(* Logix 5000 project; controller TFF vendor 1 type 14 code 107 rev 34.11; software revision 34.03; part 30 of 36 *)
(* tags used below, declared in another part *)
   Address : DINT;   // Temp Address
   Index : DINT;   // Index
   Index2 : DINT;   // Index
   ACQ002 : ALIAS FOR DigitalOutput[0];   // Emergency Stop Acknowledge
   AlarmControl : AlarmControl;   // Alarm Control
   AnalogOutput : AnalogOutput[25];   // Analog Output Array
   DigitalOutput : BOOL[256];   // Digital Output Array these bits are sent to output cards.
   FlowPath : FlowPath[64];   // Flow Path Array
   Mixer : Mixer;   // Mixer config. structure
   Options : Options;   // Options List
   PipeAnimation : PipeAnimation;   // HMI Pipe Animation Array
   PipeStatValueHMI : INT[224];   // Pipe Animation Value For HMI
   Rack_Murr_Node0_Smart : IO_Station;   // Status of Node 0 Smart
   Rack_Murr_Node1_TF2S : IO_Station;   // Status of Node 1 TF2S
   Rack_Murr_Node1_TF3S : IO_Station;   // Status of Node 1 TF3S
   Rack_Murr_Node3_PUMP : IO_Station;   // Status of Node 3 Pump
   Rack_Murr_Node4_Instrum_TFF1 : IO_Station;   // Status of Node 4 Instrum TFF1
   Rack_Murr_Node4_Instrum_TFF3 : IO_Station;   // Status of Node 4 Instrum TFF3
   Rack_Murr_Node4_Instrum_TFF5 : IO_Station;   // Status of Node 4 Instrum TFF5
   Rack_Murr_Node5_Tank100 : IO_Station;   // Status of Node 5 Tank 100L
   Rack_Murr_Node5_Tank250 : IO_Station;   // Status of Node 5 Tank 250L
   Rack_Murr_Node5_Tank50 : IO_Station;   // Status of Node 5 Tank 50L
   SIC001 : ALIAS FOR Drive[1];   // Feed Pump
   SIC001_AO : ALIAS FOR AnalogOutput[2];   // Feed Pump Speed Setpoint
   SIC002 : ALIAS FOR Drive[2];   // Transfer Pump
   SIC002_AO : ALIAS FOR AnalogOutput[3];   // Transfer Pump Speed Setpoint
   SIC003 : ALIAS FOR Drive[3];   // Mixer
   SIC003_AO : ALIAS FOR AnalogOutput[4];   // Mixer Speed Setpoint
   SysControl : SysControl;   // General system status and command
   Tank : TankManagement;   // Tank Management
   ThisSystem : SystemType;
   Valve : Valve[100];   // Valve Array
   ValveControl : ValveControl;   // Valve Control
   XC102_3 : ALIAS FOR DigitalOutput[5];   // UV Auto Zero
   XV001 : ALIAS FOR Valve[0];   // XV001
   XV002 : ALIAS FOR Valve[1];   // XV002
   XV003 : ALIAS FOR Valve[2];   // XV003
   XV004 : ALIAS FOR Valve[3];   // XV004
   XV005 : ALIAS FOR Valve[4];   // XV005
   XV006 : ALIAS FOR Valve[19];
   XV007 : ALIAS FOR Valve[20];
   XV102 : ALIAS FOR Valve[5];   // XV102
   XV401 : ALIAS FOR Valve[6];   // XV401
   XV402 : ALIAS FOR Valve[7];   // XV402
   XV403 : ALIAS FOR Valve[15];
   XV404 : ALIAS FOR Valve[16];
   XV405 : ALIAS FOR Valve[17];
   XV406 : ALIAS FOR Valve[18];
   XV411 : ALIAS FOR Valve[8];   // XV411
   XV421 : ALIAS FOR Valve[9];   // XV421
   XV431 : ALIAS FOR Valve[10];   // XV431
   XV441 : ALIAS FOR Valve[11];   // XV441
   XV501 : ALIAS FOR Valve[12];   // XV501
   XV502 : ALIAS FOR Valve[13];   // XV502
   XV901 : ALIAS FOR Valve[14];   // XV901
   Y500A : ALIAS FOR DigitalOutput[11];   // Unlock Clamshell
   Y500B : ALIAS FOR DigitalOutput[12];   // Lock Clamshell
   Y501A : ALIAS FOR DigitalOutput[10];   // Unlock Door
   Y501B : ALIAS FOR DigitalOutput[9];   // Lock Door
   Y502A : ALIAS FOR DigitalOutput[13];   // Unlock Clamshell in Door
   Y502B : ALIAS FOR DigitalOutput[14];   // Lock Clamshell in Door
   Y503A : ALIAS FOR DigitalOutput[15];   // Connect Clamshell
   Y503B : ALIAS FOR DigitalOutput[16];   // Disconnect Clamshell
(* Process, continued *)

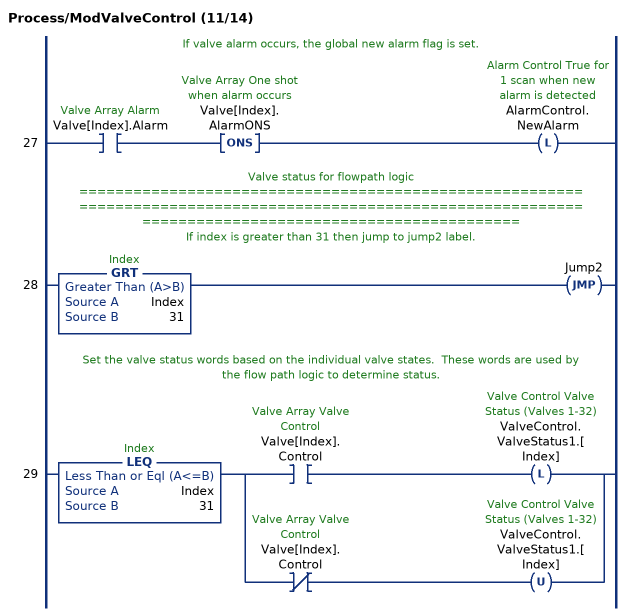
   [picture p346: Process/ModValveControl rungs 27-29]
   // If valve alarm occurs, the global new alarm flag is set.
   27: XIC(Valve[Index].Alarm)ONS(Valve[Index].AlarmONS)OTL(AlarmControl.NewAlarm);
   // Valve status for flowpath logic
   // ==========================================================================================================================================================
   // If index is greater than 31 then jump to jump2 label.
   28: GRT(Index,31)JMP(Jump2);
   // Set the valve status words based on the individual valve states.  These words are used by the flow path logic to determine status.
   29: LEQ(Index,31)[XIC(Valve[Index].Control) OTL(ValveControl.ValveStatus1.[Index]) ,XIO(Valve[Index].Control) OTU(ValveControl.ValveStatus1.[Index]) ];
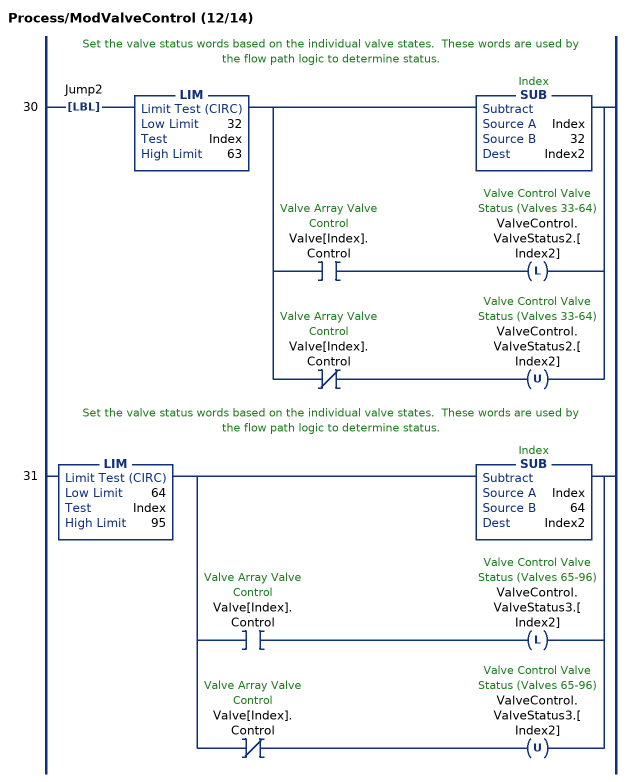
   // Set the valve status words based on the individual valve states.  These words are used by the flow path logic to determine status.
   30: LBL(Jump2)LIM(32,Index,63)[SUB(Index,32,Index2) ,XIC(Valve[Index].Control) OTL(ValveControl.ValveStatus2.[Index2]) ,XIO(Valve[Index].Control) OTU(ValveControl.ValveStatus2.[Index2]) ];
   // Set the valve status words based on the individual valve states.  These words are used by the flow path logic to determine status.
   31: LIM(64,Index,95)[SUB(Index,64,Index2) ,XIC(Valve[Index].Control) OTL(ValveControl.ValveStatus3.[Index2]) ,XIO(Valve[Index].Control) OTU(ValveControl.ValveStatus3.[Index2]) ];
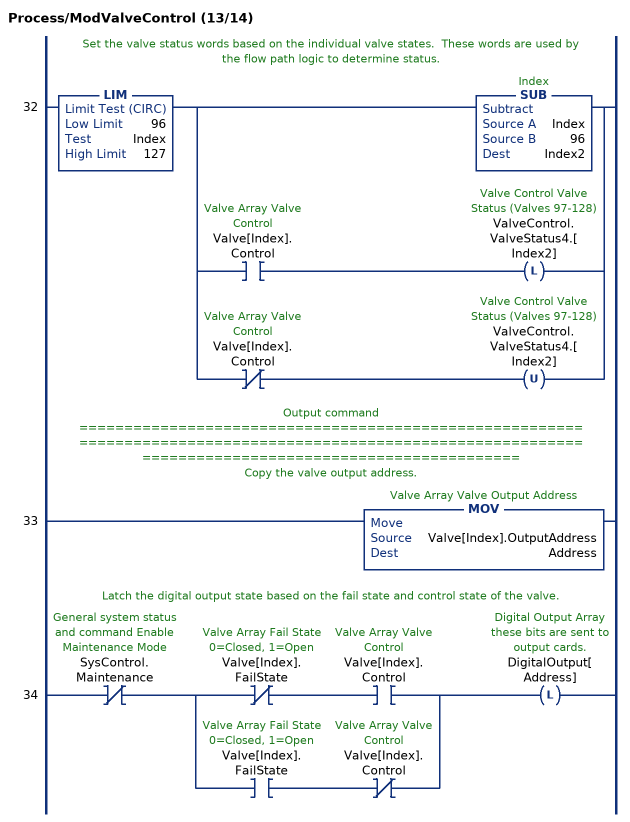
   // Set the valve status words based on the individual valve states.  These words are used by the flow path logic to determine status.
   32: LIM(96,Index,127)[SUB(Index,96,Index2) ,XIC(Valve[Index].Control) OTL(ValveControl.ValveStatus4.[Index2]) ,XIO(Valve[Index].Control) OTU(ValveControl.ValveStatus4.[Index2]) ];
   // Output command
   // ==========================================================================================================================================================
   // Copy the valve output address.
   33: MOV(Valve[Index].OutputAddress,Address);
   // Latch the digital output state based on the fail state and control state of the valve.
   34: XIO(SysControl.Maintenance)[XIO(Valve[Index].FailState) XIC(Valve[Index].Control) ,XIC(Valve[Index].FailState) XIO(Valve[Index].Control) ]OTL(DigitalOutput[Address]);
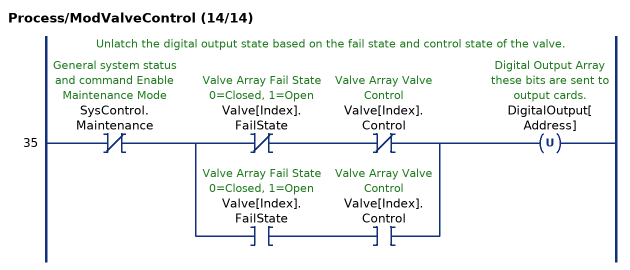
   // Unlatch the digital output state based on the fail state and control state of the valve.
   35: XIO(SysControl.Maintenance)[XIO(Valve[Index].FailState) XIO(Valve[Index].Control) ,XIC(Valve[Index].FailState) XIC(Valve[Index].Control) ]OTU(DigitalOutput[Address]);
END_ROUTINE

ROUTINE OutputAnalogPoint   (* ladder *)
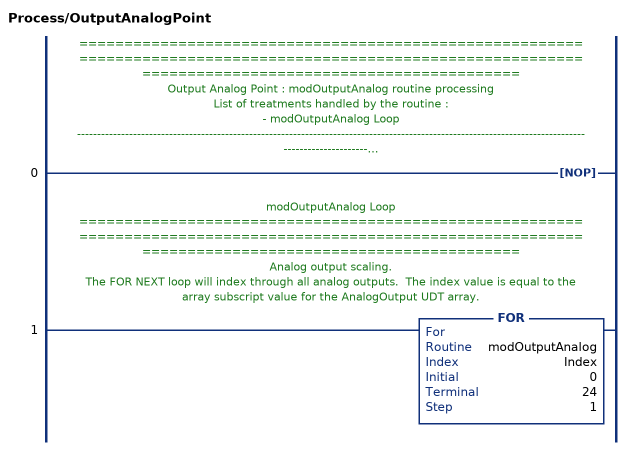
   // ==========================================================================================================================================================
   //                                                                                                             Output Analog Point : modOutputAnalog routine processing
   //                                                     List of treatments handled by the routine :
   //                                                          - modOutputAnalog Loop
   //                                                     -----------------------------------------------------------------------------------------------------------------------------------------------------
   //                                                     History
   //                                                          2019-AUG-13 - Actemium - B. Roch - Initial version for Candidate Release 3.00.00.00.a
   // ==========================================================================================================================================================
   0: NOP();
   // modOutputAnalog Loop
   // ==========================================================================================================================================================
   // Analog output scaling.
   // The FOR NEXT loop will index through all analog outputs.  The index value is equal to the array subscript value for the AnalogOutput UDT array.
   1: FOR(modOutputAnalog,Index,0,24,1);
END_ROUTINE

ROUTINE OutputAnalogRaw   (* ladder *)
// Output Routine
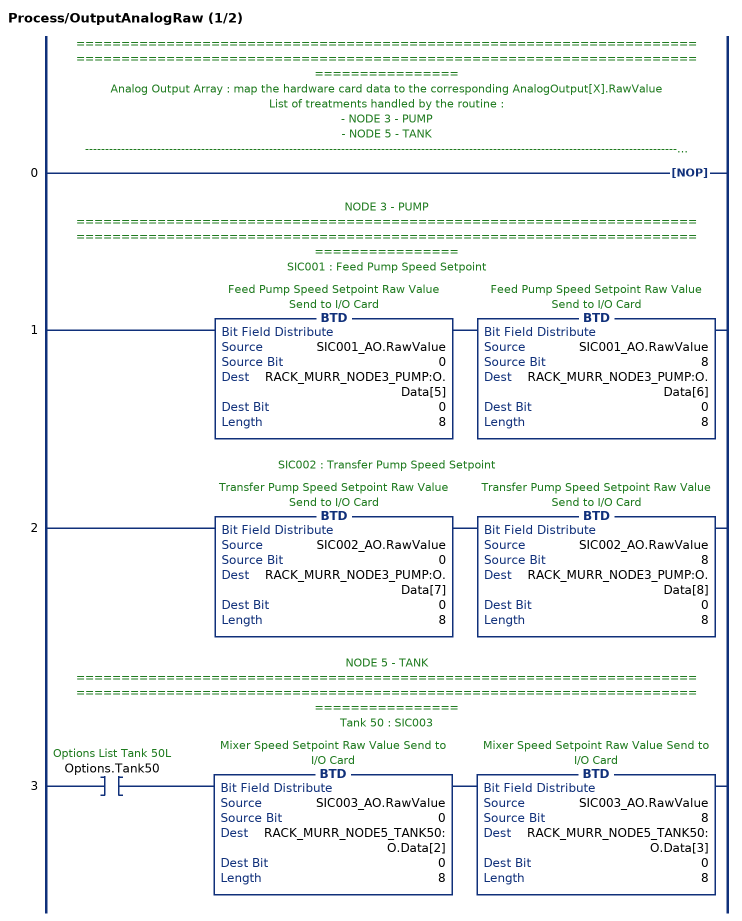
   // ==========================================================================================================================================================
   //                                                                                    Analog Output Array : map the hardware card data to the corresponding AnalogOutput[X].RawValue
   //                                                     List of treatments handled by the routine :
   //                                                   - NODE 3 - PUMP
   //                                                   - NODE 5 - TANK
   //                                                     -----------------------------------------------------------------------------------------------------------------------------------------------------
   //                                                     History
   //                                                          2019-AUG-13 - Actemium - B. Roch - Initial version for Candidate Release 3.00.00.00.a
   // ==========================================================================================================================================================
   0: NOP();
   // NODE 3 - PUMP
   // ==========================================================================================================================================================
   // SIC001 : Feed Pump Speed Setpoint
   1: BTD(SIC001_AO.RawValue,0,RACK_MURR_NODE3_PUMP:O.Data[5],0,8)BTD(SIC001_AO.RawValue,8,RACK_MURR_NODE3_PUMP:O.Data[6],0,8);
   // SIC002 : Transfer Pump Speed Setpoint
   2: BTD(SIC002_AO.RawValue,0,RACK_MURR_NODE3_PUMP:O.Data[7],0,8)BTD(SIC002_AO.RawValue,8,RACK_MURR_NODE3_PUMP:O.Data[8],0,8);
   // NODE 5 - TANK
   // ==========================================================================================================================================================
   // Tank 50 : SIC003
   3: XIC(Options.Tank50)BTD(SIC003_AO.RawValue,0,RACK_MURR_NODE5_TANK50:O.Data[2],0,8)BTD(SIC003_AO.RawValue,8,RACK_MURR_NODE5_TANK50:O.Data[3],0,8);
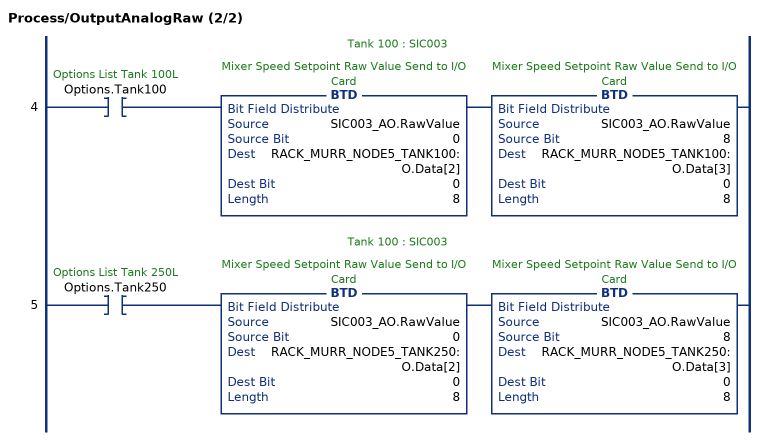
   // Tank 100 : SIC003
   4: XIC(Options.Tank100)BTD(SIC003_AO.RawValue,0,RACK_MURR_NODE5_TANK100:O.Data[2],0,8)BTD(SIC003_AO.RawValue,8,RACK_MURR_NODE5_TANK100:O.Data[3],0,8);
   // Tank 100 : SIC003
   5: XIC(Options.Tank250)BTD(SIC003_AO.RawValue,0,RACK_MURR_NODE5_TANK250:O.Data[2],0,8)BTD(SIC003_AO.RawValue,8,RACK_MURR_NODE5_TANK250:O.Data[3],0,8);
END_ROUTINE

ROUTINE OutputDigitalRaw   (* ladder *)
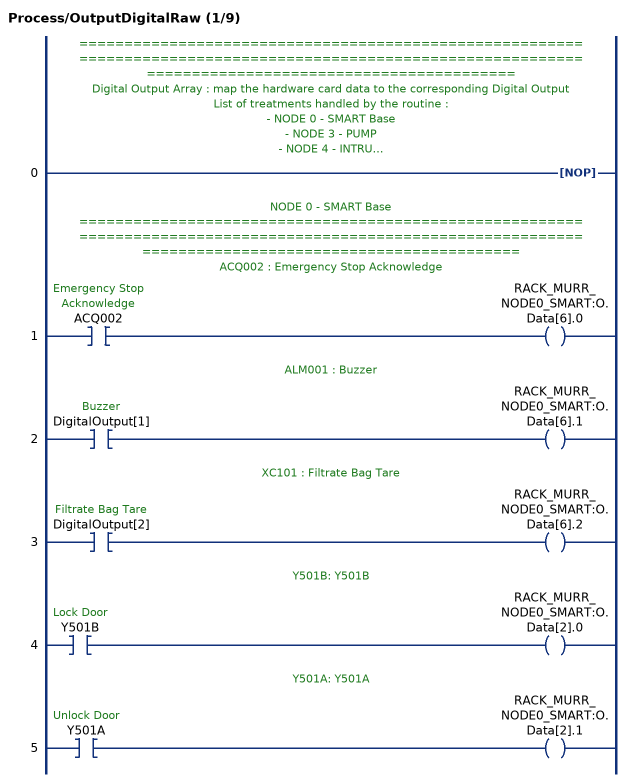
   // =========================================================================================================================================================
   //                                                                                          Digital Output Array : map the hardware card data to the corresponding Digital Output
   //                                                     List of treatments handled by the routine :
   //                                                    - NODE 0 - SMART Base
   //                                                    - NODE 3 - PUMP
   //                                                    - NODE 4 - INTRUM
   //                                                    - NODE 5 - TANK
   //                                                    - NODE 1 - TF2S
   //                                                    - NODE 1 - TF3S
   //                                                     -----------------------------------------------------------------------------------------------------------------------------------------------------
   //                                                     History
   //                    2019-AUG-13 - Actemium - B. Roch - Initial version for Candidate Release 3.00.00.00.a
   // 	2019-SEP-16 - ACTEMIUM - Q. Spindler - Modifications for Candidate Release 3.00.00.00.c
   // 					- Change mapping IO for Inlets valves
   // 	2021-APR-13 - DAVIDSON- Ch. ARBOGAST - Modifications for Candidate Release 3.01.00.00.a
   // 			Add rungs 20 to 25: output valves XV403-404-405-406-006-007
   // ==========================================================================================================================================================
   0: NOP();
   // NODE 0 - SMART Base
   // ==========================================================================================================================================================
   // ACQ002 : Emergency Stop Acknowledge
   1: XIC(ACQ002)OTE(RACK_MURR_NODE0_SMART:O.Data[6].0);
   // ALM001 : Buzzer
   2: XIC(DigitalOutput[1])OTE(RACK_MURR_NODE0_SMART:O.Data[6].1);
   // XC101 : Filtrate Bag Tare
   3: XIC(DigitalOutput[2])OTE(RACK_MURR_NODE0_SMART:O.Data[6].2);
   // Y501B: Y501B
   4: XIC(Y501B)OTE(RACK_MURR_NODE0_SMART:O.Data[2].0);
   // Y501A: Y501A
   5: XIC(Y501A)OTE(RACK_MURR_NODE0_SMART:O.Data[2].1);
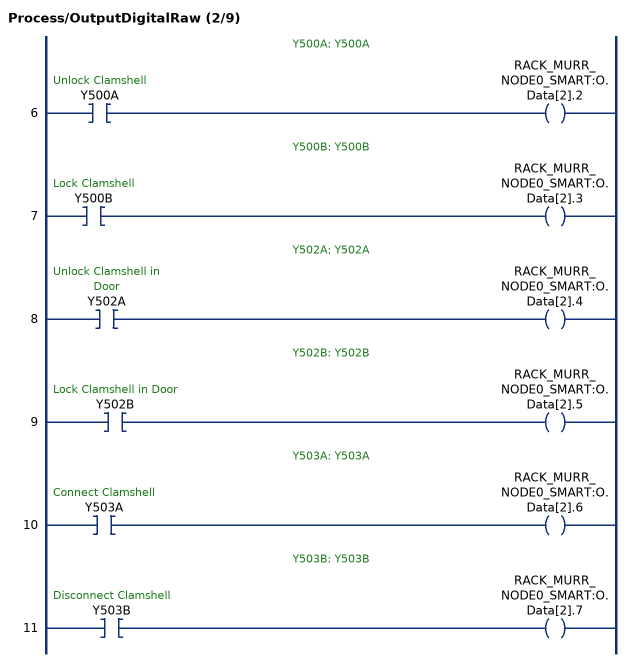
   // Y500A: Y500A
   6: XIC(Y500A)OTE(RACK_MURR_NODE0_SMART:O.Data[2].2);
   // Y500B: Y500B
   7: XIC(Y500B)OTE(RACK_MURR_NODE0_SMART:O.Data[2].3);
   // Y502A: Y502A
   8: XIC(Y502A)OTE(RACK_MURR_NODE0_SMART:O.Data[2].4);
   // Y502B: Y502B
   9: XIC(Y502B)OTE(RACK_MURR_NODE0_SMART:O.Data[2].5);
   // Y503A: Y503A
   10: XIC(Y503A)OTE(RACK_MURR_NODE0_SMART:O.Data[2].6);
   // Y503B: Y503B
   11: XIC(Y503B)OTE(RACK_MURR_NODE0_SMART:O.Data[2].7);
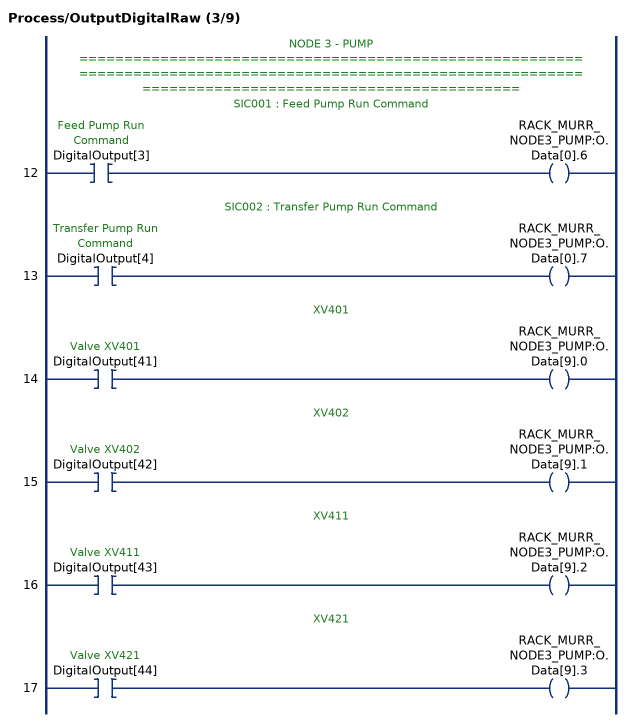
   // NODE 3 - PUMP
   // ==========================================================================================================================================================
   // SIC001 : Feed Pump Run Command
   12: XIC(DigitalOutput[3])OTE(RACK_MURR_NODE3_PUMP:O.Data[0].6);
   // SIC002 : Transfer Pump Run Command
   13: XIC(DigitalOutput[4])OTE(RACK_MURR_NODE3_PUMP:O.Data[0].7);
   // XV401
   14: XIC(DigitalOutput[41])OTE(RACK_MURR_NODE3_PUMP:O.Data[9].0);
   // XV402
   15: XIC(DigitalOutput[42])OTE(RACK_MURR_NODE3_PUMP:O.Data[9].1);
   // XV411
   16: XIC(DigitalOutput[43])OTE(RACK_MURR_NODE3_PUMP:O.Data[9].2);
   // XV421
   17: XIC(DigitalOutput[44])OTE(RACK_MURR_NODE3_PUMP:O.Data[9].3);
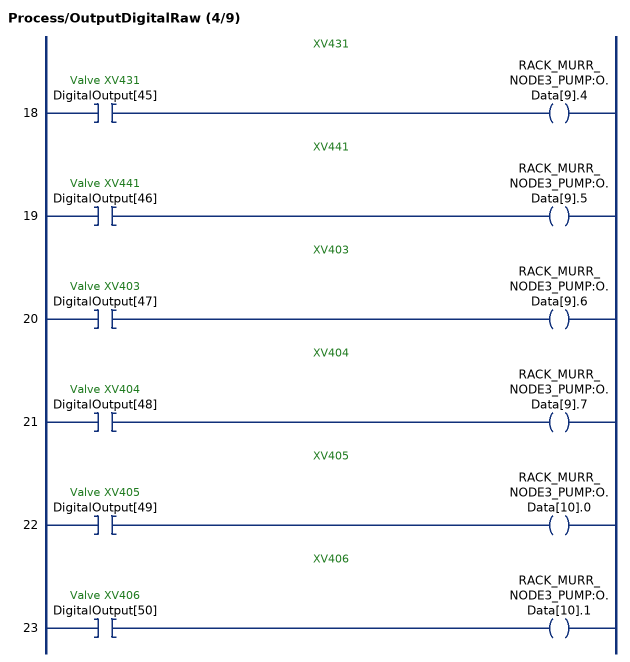
   // XV431
   18: XIC(DigitalOutput[45])OTE(RACK_MURR_NODE3_PUMP:O.Data[9].4);
   // XV441
   19: XIC(DigitalOutput[46])OTE(RACK_MURR_NODE3_PUMP:O.Data[9].5);
   // XV403
   20: XIC(DigitalOutput[47])OTE(RACK_MURR_NODE3_PUMP:O.Data[9].6);
   // XV404
   21: XIC(DigitalOutput[48])OTE(RACK_MURR_NODE3_PUMP:O.Data[9].7);
   // XV405
   22: XIC(DigitalOutput[49])OTE(RACK_MURR_NODE3_PUMP:O.Data[10].0);
   // XV406
   23: XIC(DigitalOutput[50])OTE(RACK_MURR_NODE3_PUMP:O.Data[10].1);
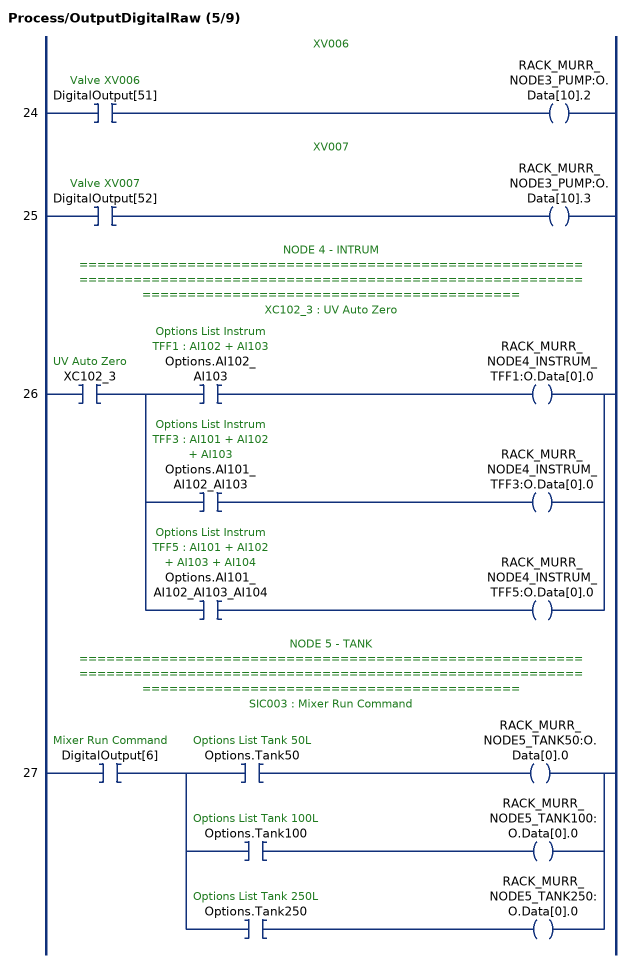
   // XV006
   24: XIC(DigitalOutput[51])OTE(RACK_MURR_NODE3_PUMP:O.Data[10].2);
   // XV007
   25: XIC(DigitalOutput[52])OTE(RACK_MURR_NODE3_PUMP:O.Data[10].3);
   // NODE 4 - INTRUM
   // ==========================================================================================================================================================
   // XC102_3 : UV Auto Zero
   26: XIC(XC102_3)[XIC(Options.AI102_AI103) OTE(RACK_MURR_NODE4_INSTRUM_TFF1:O.Data[0].0) ,XIC(Options.AI101_AI102_AI103) OTE(RACK_MURR_NODE4_INSTRUM_TFF3:O.Data[0].0) ,XIC(Options.AI101_AI102_AI103_AI104) OTE(RACK_MURR_NODE4_INSTRUM_TFF5:O.Data[0].0) ];
   // NODE 5 - TANK
   // ==========================================================================================================================================================
   // SIC003 : Mixer Run Command
   27: XIC(DigitalOutput[6])[XIC(Options.Tank50) OTE(RACK_MURR_NODE5_TANK50:O.Data[0].0) ,XIC(Options.Tank100) OTE(RACK_MURR_NODE5_TANK100:O.Data[0].0) ,XIC(Options.Tank250) OTE(RACK_MURR_NODE5_TANK250:O.Data[0].0) ];
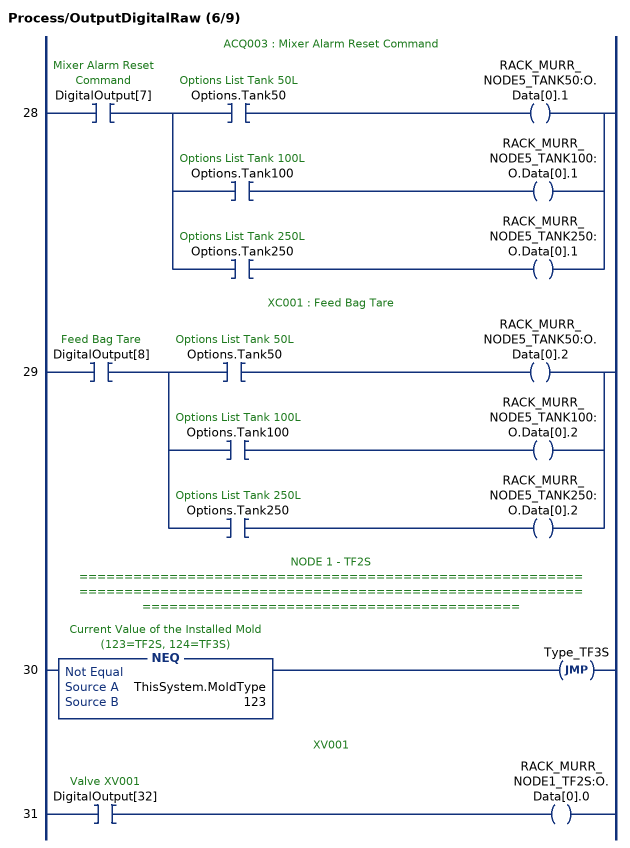
   // ACQ003 : Mixer Alarm Reset Command
   28: XIC(DigitalOutput[7])[XIC(Options.Tank50) OTE(RACK_MURR_NODE5_TANK50:O.Data[0].1) ,XIC(Options.Tank100) OTE(RACK_MURR_NODE5_TANK100:O.Data[0].1) ,XIC(Options.Tank250) OTE(RACK_MURR_NODE5_TANK250:O.Data[0].1) ];
   // XC001 : Feed Bag Tare
   29: XIC(DigitalOutput[8])[XIC(Options.Tank50) OTE(RACK_MURR_NODE5_TANK50:O.Data[0].2) ,XIC(Options.Tank100) OTE(RACK_MURR_NODE5_TANK100:O.Data[0].2) ,XIC(Options.Tank250) OTE(RACK_MURR_NODE5_TANK250:O.Data[0].2) ];
   // NODE 1 - TF2S
   // ==========================================================================================================================================================
   30: NEQ(ThisSystem.MoldType,123)JMP(Type_TF3S);
   // XV001
   31: XIC(DigitalOutput[32])OTE(RACK_MURR_NODE1_TF2S:O.Data[0].0);
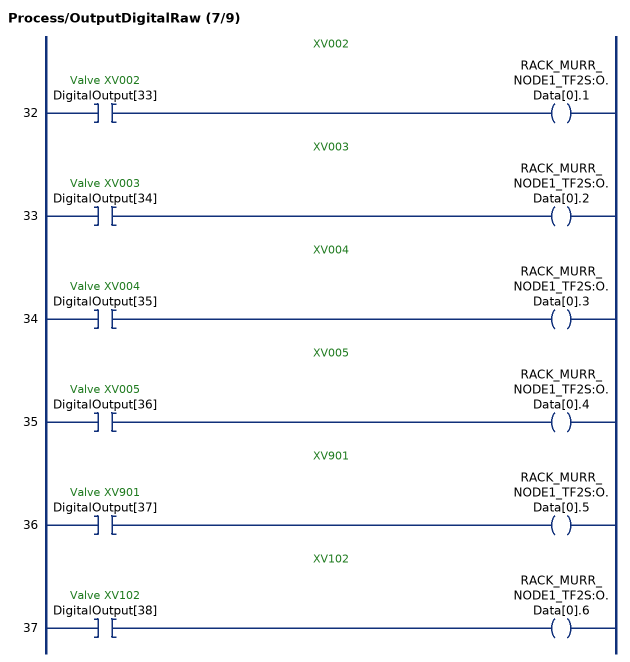
   // XV002
   32: XIC(DigitalOutput[33])OTE(RACK_MURR_NODE1_TF2S:O.Data[0].1);
   // XV003
   33: XIC(DigitalOutput[34])OTE(RACK_MURR_NODE1_TF2S:O.Data[0].2);
   // XV004
   34: XIC(DigitalOutput[35])OTE(RACK_MURR_NODE1_TF2S:O.Data[0].3);
   // XV005
   35: XIC(DigitalOutput[36])OTE(RACK_MURR_NODE1_TF2S:O.Data[0].4);
   // XV901
   36: XIC(DigitalOutput[37])OTE(RACK_MURR_NODE1_TF2S:O.Data[0].5);
   // XV102
   37: XIC(DigitalOutput[38])OTE(RACK_MURR_NODE1_TF2S:O.Data[0].6);
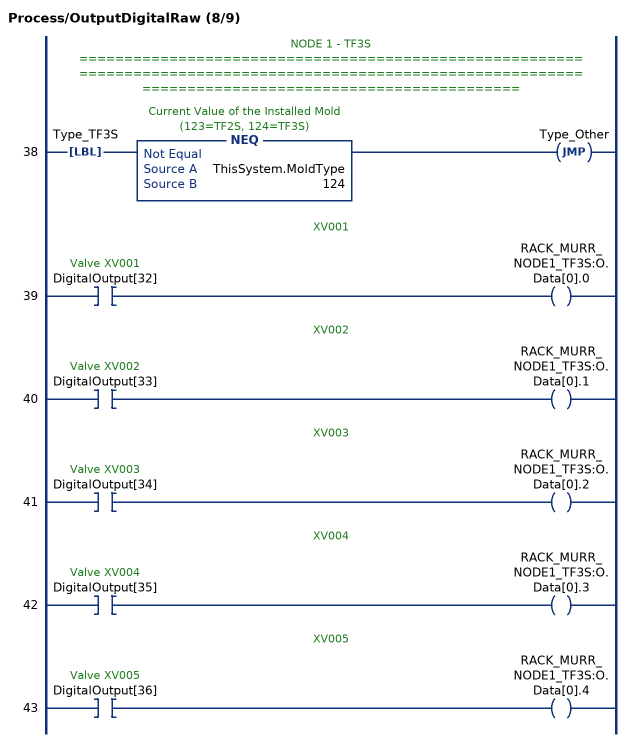
   // NODE 1 - TF3S
   // ==========================================================================================================================================================
   38: LBL(Type_TF3S)NEQ(ThisSystem.MoldType,124)JMP(Type_Other);
   // XV001
   39: XIC(DigitalOutput[32])OTE(RACK_MURR_NODE1_TF3S:O.Data[0].0);
   // XV002
   40: XIC(DigitalOutput[33])OTE(RACK_MURR_NODE1_TF3S:O.Data[0].1);
   // XV003
   41: XIC(DigitalOutput[34])OTE(RACK_MURR_NODE1_TF3S:O.Data[0].2);
   // XV004
   42: XIC(DigitalOutput[35])OTE(RACK_MURR_NODE1_TF3S:O.Data[0].3);
   // XV005
   43: XIC(DigitalOutput[36])OTE(RACK_MURR_NODE1_TF3S:O.Data[0].4);
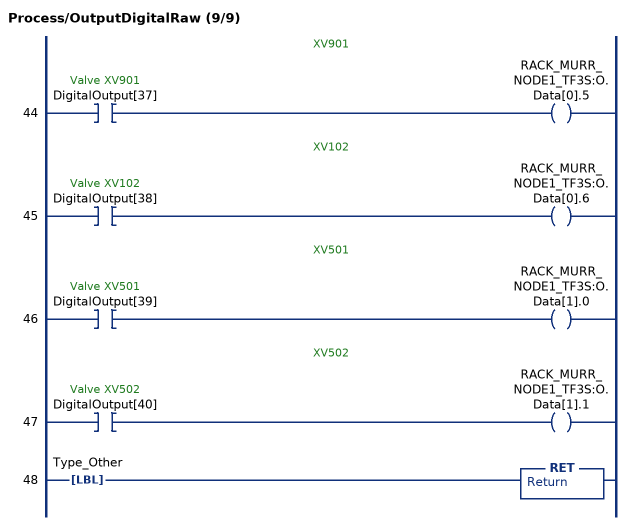
   // XV901
   44: XIC(DigitalOutput[37])OTE(RACK_MURR_NODE1_TF3S:O.Data[0].5);
   // XV102
   45: XIC(DigitalOutput[38])OTE(RACK_MURR_NODE1_TF3S:O.Data[0].6);
   // XV501
   46: XIC(DigitalOutput[39])OTE(RACK_MURR_NODE1_TF3S:O.Data[1].0);
   // XV502
   47: XIC(DigitalOutput[40])OTE(RACK_MURR_NODE1_TF3S:O.Data[1].1);
   48: LBL(Type_Other)RET();
END_ROUTINE

ROUTINE OutputProcessing   (* ladder *)
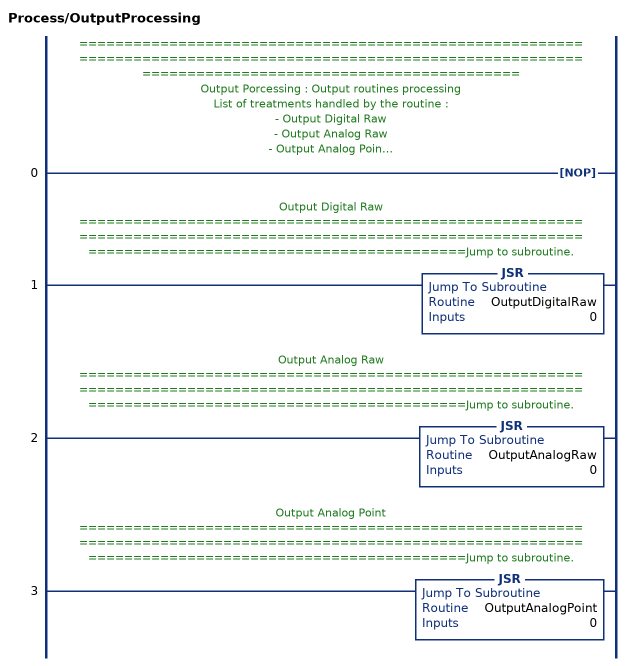
   // ==========================================================================================================================================================
   //                                                                                                                  Output Porcessing : Output routines processing
   //                                                     List of treatments handled by the routine :
   //                                                          - Output Digital Raw
   //                                                          - Output Analog Raw
   //                                                          - Output Analog Point
   //                                                     -----------------------------------------------------------------------------------------------------------------------------------------------------
   //                                                     History
   //                                                          2019-AUG-13 - Actemium - B. Roch - Initial version for Candidate Release 3.00.00.00.a
   // ==========================================================================================================================================================
   0: NOP();
   // Output Digital Raw
   // ==========================================================================================================================================================Jump to subroutine.
   1: JSR(OutputDigitalRaw,0);
   // Output Analog Raw
   // ==========================================================================================================================================================Jump to subroutine.
   2: JSR(OutputAnalogRaw,0);
   // Output Analog Point
   // ==========================================================================================================================================================Jump to subroutine.
   3: JSR(OutputAnalogPoint,0);
END_ROUTINE

ROUTINE PipeAnimation   (* ladder *)
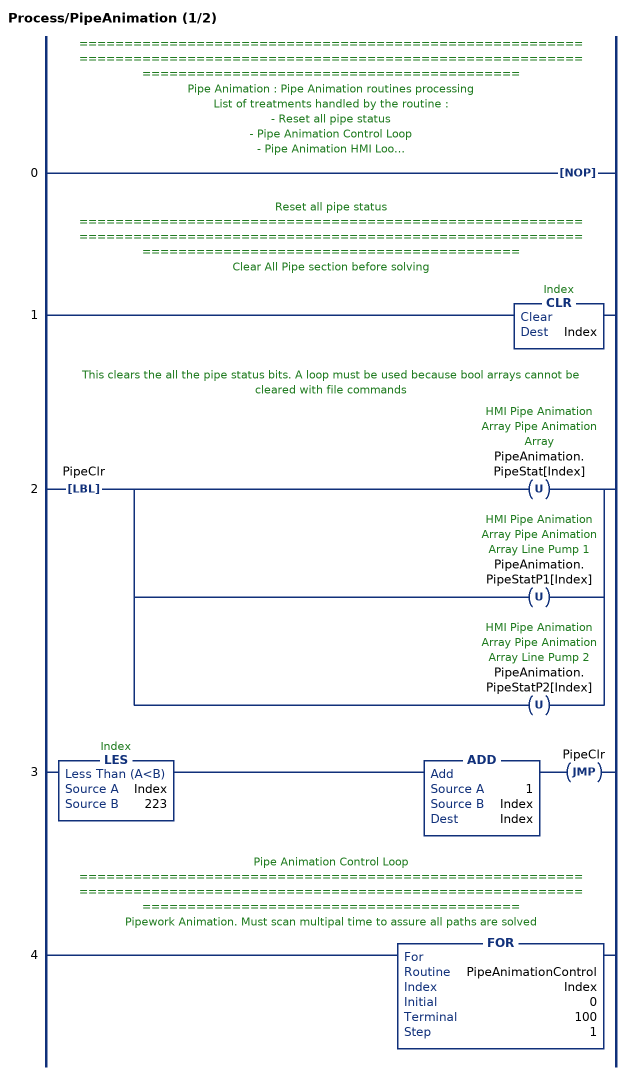
   // ==========================================================================================================================================================
   //                                                                                                               Pipe Animation : Pipe Animation routines processing
   //                                                     List of treatments handled by the routine :
   //                                                          - Reset all pipe status
   //                                                          - Pipe Animation Control Loop
   //                                                          - Pipe Animation HMI Loop
   //                                                     -----------------------------------------------------------------------------------------------------------------------------------------------------
   //                                                     History
   //                                                         2019-AUG-13 - Actemium - B. Roch - Initial version for Candidate Release 3.00.00.00.a
   // ==========================================================================================================================================================
   0: NOP();
   // Reset all pipe status
   // ==========================================================================================================================================================
   // Clear All Pipe section before solving
   1: CLR(Index);
   // This clears the all the pipe status bits. A loop must be used because bool arrays cannot be cleared with file commands
   2: LBL(PipeClr)[OTU(PipeAnimation.PipeStat[Index]) ,OTU(PipeAnimation.PipeStatP1[Index]) ,OTU(PipeAnimation.PipeStatP2[Index]) ];
   3: LES(Index,223)ADD(1,Index,Index)JMP(PipeClr);
   // Pipe Animation Control Loop
   // ==========================================================================================================================================================
   // Pipework Animation. Must scan multipal time to assure all paths are solved
   4: FOR(PipeAnimationControl,Index,0,100,1);
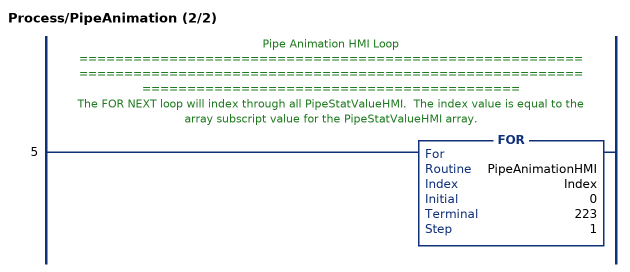
   // Pipe Animation HMI Loop
   // ==========================================================================================================================================================
   // The FOR NEXT loop will index through all PipeStatValueHMI.  The index value is equal to the array subscript value for the PipeStatValueHMI array.
   5: FOR(PipeAnimationHMI,Index,0,223,1);
END_ROUTINE
